FUNCTION_BLOCK RecoveryTarget (* Valid target for importer recovery *)
  (* Standard: 61499-1; Description: Copyright (c) 2026 Martin Erich Jobst This program and the accompanying materials are made available under the terms of the Eclipse Public License 2.0 which is available at https://www.eclipse.org/legal/epl-2.0/ SPDX-License-Identifier: EPL-2.0 *)
  (* Version 1.0, 2026-10-23, Martin Jobst *)
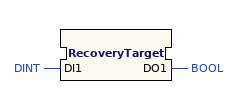
  VAR_INPUT
    DI1 : DINT;
  END_VAR
  VAR_OUTPUT
    DO1 : BOOL;
  END_VAR
END_FUNCTION_BLOCK
